(* IEC 61131-3 sources: dummvinci-rosetta-plc/src/plc_mcp/library/patterns, 6 files *)

(* ---- FB_AlarmManager.st ---- *)
(* =====================================================================
   FB_AlarmManager — aggregate N alarm points (IEC 62682 / ISA-18.2)
   dummvinci-rosetta-plc engineering library

   Aggregates the OUTPUT arrays of FB_AlarmPoint instances: per-class
   counts, unacked count, horn drive, and FIRST-OUT capture (which alarm
   started the trip cascade — the question every breakdown review asks).

   USAGE
     The application owns the FB_AlarmPoint instances and copies their
     outputs into the three arrays each cycle (or maps them directly):
       aActive[i]  := fbAlm_i.xActive;
       aUnacked[i] := fbAlm_i.xUnacked;
       aClass[i]   := fbAlm_i.eClass;
     then calls:
       fbMgr(nPoints := <used>, aActive := ..., aUnacked := ..., aClass := ...);
     Group acknowledge: wire fbMgr.xAckPulse into every point's xAck.
     Sizing: ARRAY[1..64] here — adjust bound + nPoints per project.

   DISCLAIMER — draft engineering input, review + FAT mandatory.
   NOT for safety-instrumented functions (SAFETY.md / H11).
   ===================================================================== *)

FUNCTION_BLOCK FB_AlarmManager
VAR_INPUT
    nPoints    : INT;    (* number of points actually used, <= 64 *)
    xGroupAck  : BOOL;   (* operator group-acknowledge command    *)
    xHornReset : BOOL;   (* silence horn without acknowledging    *)
END_VAR
VAR_IN_OUT
    aActive  : ARRAY[1..64] OF BOOL;
    aUnacked : ARRAY[1..64] OF BOOL;
    aClass   : ARRAY[1..64] OF INT;   (* 2 FAULT / 1 WARNING / 0 EVENT *)
END_VAR
VAR_OUTPUT
    nActive        : INT;
    nUnacked       : INT;
    nActiveFault   : INT;
    nActiveWarning : INT;
    iFirstOut      : INT;    (* index of first-out alarm, 0 = none *)
    xHorn          : BOOL;   (* unacked FAULT/WARNING present      *)
    xAckPulse      : BOOL;   (* wire into every point's xAck input *)
END_VAR
VAR
    i           : INT;
    aPrevActive : ARRAY[1..64] OF BOOL;
    nPrevActive : INT;
    xHornMuted  : BOOL;
    trigAck     : R_TRIG;
END_VAR

trigAck(CLK := xGroupAck);
xAckPulse := trigAck.Q;

nActive := 0;
nUnacked := 0;
nActiveFault := 0;
nActiveWarning := 0;

FOR i := 1 TO nPoints DO
    IF aActive[i] THEN
        nActive := nActive + 1;
        IF aClass[i] = 2 THEN
            nActiveFault := nActiveFault + 1;
        END_IF;
        IF aClass[i] = 1 THEN
            nActiveWarning := nActiveWarning + 1;
        END_IF;
    END_IF;
    IF aUnacked[i] THEN
        nUnacked := nUnacked + 1;
    END_IF;

    (* first-out: the point that went active while nothing was active *)
    IF aActive[i] AND NOT aPrevActive[i]
       AND (nPrevActive = 0) AND (iFirstOut = 0) THEN
        iFirstOut := i;
    END_IF;
    aPrevActive[i] := aActive[i];
END_FOR;

(* first-out clears only when the plant is alarm-free again *)
IF nActive = 0 THEN
    iFirstOut := 0;
END_IF;
nPrevActive := nActive;

(* horn: any unacked FAULT/WARNING; mute survives until all acked *)
IF xHornReset THEN
    xHornMuted := TRUE;
END_IF;
IF nUnacked = 0 THEN
    xHornMuted := FALSE;
END_IF;
xHorn := (nUnacked > 0) AND NOT xHornMuted;

END_FUNCTION_BLOCK

(* ---- FB_AlarmPoint.st ---- *)
(* =====================================================================
   FB_AlarmPoint — single alarm point state machine
   dummvinci-rosetta-plc engineering library

   STANDARD BASIS
     IEC 62682 / ISA-18.2 alarm states:
       0 = NORM        normal, inactive
       1 = UNACK_ALM   active, unacknowledged
       2 = ACK_ALM     active, acknowledged
       3 = UNACK_RTN   returned to normal, still unacknowledged
     Meldeklassen mapping (German practice):
       eClass 2 = FAULT   (Störung)   — trips/stops the function
       eClass 1 = WARNING (Warnung)   — degraded, action required
       eClass 0 = EVENT   (Meldung)   — information, logged only

   USAGE
     One instance per alarm point. Call every task cycle:
       fbAlm(xIn := <raw condition>, xAck := <ack cmd>, xReset := <reset>);
     Wire xAppeared/xDisappeared/xAckEdge into FB_EventLogger for the
     historian, and xActive/xUnacked/eClass arrays into FB_AlarmManager.

   DISCLAIMER — draft engineering input, review + FAT mandatory.
   NOT for safety-instrumented functions (see SAFETY.md / H11): e-stop,
   overload, interlock chains belong on a certified safety CPU.
   ===================================================================== *)

FUNCTION_BLOCK FB_AlarmPoint
VAR_INPUT
    xIn        : BOOL;   (* raw alarm condition, TRUE = abnormal *)
    xAck       : BOOL;   (* acknowledge command (operator/group)  *)
    xReset     : BOOL;   (* reset for latched alarms              *)
    xLatching  : BOOL;   (* TRUE: stays active until xReset       *)
    tOnDelay   : TIME;   (* debounce before alarm becomes active  *)
    tOffDelay  : TIME;   (* delay before return-to-normal         *)
    iPriority  : INT;    (* 1=low .. 4=critical (per philosophy)  *)
    eClass     : INT;    (* 2=FAULT, 1=WARNING, 0=EVENT           *)
    diCode     : DINT;   (* error code for catalog/historian      *)
END_VAR
VAR_OUTPUT
    xActive       : BOOL;  (* alarm condition present (qualified) *)
    xUnacked      : BOOL;  (* requires operator acknowledgement   *)
    eState        : INT;   (* 0 NORM / 1 UNACK_ALM / 2 ACK_ALM / 3 UNACK_RTN *)
    xAppeared     : BOOL;  (* one-cycle pulse: alarm appeared     *)
    xDisappeared  : BOOL;  (* one-cycle pulse: alarm cleared      *)
    xAckEdge      : BOOL;  (* one-cycle pulse: acknowledged       *)
END_VAR
VAR
    tonQualify  : TON;
    tonClear    : TON;
    xQualified  : BOOL;
    xLatched    : BOOL;
    trigApp     : R_TRIG;
    trigDis     : F_TRIG;
    trigAck     : R_TRIG;
END_VAR

(* --- qualification: debounce both directions ---------------------- *)
tonQualify(IN := xIn, PT := tOnDelay);
tonClear(IN := NOT xIn, PT := tOffDelay);

IF tonQualify.Q THEN
    xQualified := TRUE;
END_IF;
IF tonClear.Q THEN
    xQualified := FALSE;
END_IF;

(* --- latching ------------------------------------------------------ *)
IF xLatching AND xQualified THEN
    xLatched := TRUE;
END_IF;
IF xReset AND NOT xQualified THEN
    xLatched := FALSE;
END_IF;

xActive := xQualified OR (xLatching AND xLatched);

(* --- ack edge: evaluate BEFORE the state machine clears xUnacked --- *)
trigAck(CLK := xAck AND xUnacked);
xAckEdge := trigAck.Q;

(* --- IEC 62682 state machine --------------------------------------- *)
CASE eState OF
    0: (* NORM *)
        IF xActive THEN
            eState := 1;
            xUnacked := TRUE;
        END_IF;
    1: (* UNACK_ALM *)
        IF xAck THEN
            eState := 2;
            xUnacked := FALSE;
        ELSIF NOT xActive THEN
            eState := 3;
        END_IF;
    2: (* ACK_ALM *)
        IF NOT xActive THEN
            eState := 0;
        END_IF;
    3: (* UNACK_RTN *)
        IF xAck THEN
            eState := 0;
            xUnacked := FALSE;
        ELSIF xActive THEN
            eState := 1;
        END_IF;
END_CASE;

(* --- edges for the historian ---------------------------------------- *)
trigApp(CLK := xActive);
xAppeared := trigApp.Q;
trigDis(CLK := xActive);
xDisappeared := trigDis.Q;

END_FUNCTION_BLOCK

(* ---- FB_CommsWatchdog.st ---- *)
(* =====================================================================
   FB_CommsWatchdog — communication supervision (DIAGNOSTICS ONLY)
   dummvinci-rosetta-plc engineering library

   Supervises a cyclic link (Modbus TCP slave, HMI, remote I/O) via a
   heartbeat counter that the remote increments. If the counter stops
   changing for tTimeout, the link is declared down — feed that into an
   FB_AlarmPoint (class WARNING or FAULT per the alarm philosophy).

   ⚠ THIS IS NOT A SAFETY WATCHDOG. A watchdog whose timeout must bring
   the machine to a safe state is a safety function — that belongs on a
   certified safety CPU (AC500-S) per SAFETY.md / hazard H11. This block
   only *reports* link health.

   USAGE (Modbus TCP to an ACS880 example)
     Map a drive register that changes continuously (e.g. a counter or
     the actual-speed word) into diHeartbeat:
       fbWd(diHeartbeat := <mapped register>, tTimeout := T#3s);

   DISCLAIMER — draft engineering input, review + FAT mandatory.
   ===================================================================== *)

FUNCTION_BLOCK FB_CommsWatchdog
VAR_INPUT
    diHeartbeat : DINT;   (* value the remote updates cyclically *)
    tTimeout    : TIME;   (* declare down after this long unchanged *)
END_VAR
VAR_OUTPUT
    xCommsOk  : BOOL;
    xTimeout  : BOOL;
    udiDrops  : UDINT;    (* number of times the link went down *)
END_VAR
VAR
    diPrev   : DINT;
    tonStale : TON;
    trigDown : R_TRIG;
END_VAR

tonStale(IN := (diHeartbeat = diPrev), PT := tTimeout);
diPrev := diHeartbeat;

xTimeout := tonStale.Q;
xCommsOk := NOT xTimeout;

trigDown(CLK := xTimeout);
IF trigDown.Q THEN
    udiDrops := udiDrops + 1;
END_IF;

END_FUNCTION_BLOCK

(* ---- FB_DriveDiagACS880.st ---- *)
(* =====================================================================
   FB_DriveDiagACS880 — ACS880 fault/warning capture for the historian
   dummvinci-rosetta-plc engineering library

   Captures the active fault/warning codes of an ABB ACS880 drive (read
   over Modbus TCP / PROFINET) and converts them to hex strings that key
   directly into the error-code catalog (plc_errorcode_lookup, source
   "acs880") for cause + remedy.

   REGISTER MAPPING (project-specific — TODO verify against YOUR comms
   mapping in Drive Composer Pro; typical parameters):
     04.01  Tripping fault code    -> uiFaultCode
     04.06  Active warning code    -> uiWarnCode
     Status word bit FAULTED       -> xDriveFaulted
     Status word bit WARNING       -> xDriveWarning

   USAGE
     fbDiag(uiFaultCode := <mapped 04.01>, uiWarnCode := <mapped 04.06>,
            xDriveFaulted := <SW bit>, xDriveWarning := <SW bit>);
     On xNewFault: log to FB_EventLogger with diCode := fbDiag.diFaultCode
     and look the hex string up in the catalog.

   DISCLAIMER — draft engineering input, review + FAT mandatory. Codes and
   remedies come from the catalog, which must be verified against the
   ACS880 firmware manual for the installed FW revision.
   ===================================================================== *)

FUNCTION_BLOCK FB_DriveDiagACS880
VAR_INPUT
    uiFaultCode   : UINT;   (* drive par 04.01 via comms *)
    uiWarnCode    : UINT;   (* drive par 04.06 via comms *)
    xDriveFaulted : BOOL;   (* status word: faulted      *)
    xDriveWarning : BOOL;   (* status word: warning      *)
END_VAR
VAR_OUTPUT
    xFault      : BOOL;
    xWarning    : BOOL;
    diFaultCode : DINT;         (* numeric, for FB_EventLogger *)
    sFaultHex   : STRING(7);    (* catalog key, e.g. '2310'    *)
    sWarnHex    : STRING(7);
    xNewFault   : BOOL;         (* one-cycle pulse             *)
    xNewWarning : BOOL;
END_VAR
VAR
    trigF : R_TRIG;
    trigW : R_TRIG;
    uiTmp : UINT;
    iNib  : INT;
    i     : INT;
    sHex  : STRING(7);
END_VAR

xFault := xDriveFaulted;
xWarning := xDriveWarning;
diFaultCode := TO_DINT(uiFaultCode);

(* --- UINT -> 4-digit hex string (ACS880 codes read as hex) ---------
   MID signature per IEC 61131-3 / CODESYS Standard library:
   MID(IN, L, P) = L characters starting at position P (1-based).
   So MID('0123456789ABCDEF', L := 1, P := iNib + 1) extracts exactly
   ONE nibble character. Do not swap to (pos, len) — that is a
   different vendor convention. ------------------------------------- *)
sHex := '';
uiTmp := uiFaultCode;
FOR i := 1 TO 4 DO
    iNib := TO_INT(uiTmp MOD 16);
    sHex := CONCAT(MID(IN := '0123456789ABCDEF', L := 1, P := iNib + 1),
                   sHex);
    uiTmp := uiTmp / 16;
END_FOR;
sFaultHex := sHex;

sHex := '';
uiTmp := uiWarnCode;
FOR i := 1 TO 4 DO
    iNib := TO_INT(uiTmp MOD 16);
    sHex := CONCAT(MID(IN := '0123456789ABCDEF', L := 1, P := iNib + 1),
                   sHex);
    uiTmp := uiTmp / 16;
END_FOR;
sWarnHex := sHex;

trigF(CLK := xDriveFaulted);
xNewFault := trigF.Q;
trigW(CLK := xDriveWarning);
xNewWarning := trigW.Q;

END_FUNCTION_BLOCK

(* ---- FB_EventLogger.st ---- *)
(* =====================================================================
   FB_EventLogger — sequence-of-events ring-buffer historian
   dummvinci-rosetta-plc engineering library

   In-PLC SoE log: every alarm appearance/clearance/acknowledgement is
   stamped and kept in a retained ring buffer for breakdown analysis and
   HMI display. Design rationale: docs/library/HISTORIAN-DESIGN.md
   (resolution limits, time sync, when to use an external historian).

   USAGE
     One instance per log. Feed one event per rising edge of xLog —
     typically chained from FB_AlarmPoint edges:
       IF fbAlm.xAppeared THEN
           fbLog(xLog := TRUE, diCode := fbAlm.diCode,
                 eClass := fbAlm.eClass, eEdge := 0, rValue := <pv>,
                 dtNow := <rtc>, uiMsOfSec := <ms>);
       END_IF
     eEdge: 0 = APPEARED, 1 = DISAPPEARED, 2 = ACKED.
     (* TODO platform binding: dtNow/uiMsOfSec must come from the CPU RTC
        — e.g. AC500 V3 SysTimeRtc / DT clock FBs. Timestamp AT SOURCE,
        in the same task that detects the edge. *)
     Buffer: ARRAY[0..255] here — size per project; RETAIN memory is a
     real CPU budget, verify against the CPU's retain capacity.

   TYPES (move to a DUT object on Automation Builder import)
   ===================================================================== *)

TYPE ST_Event :
STRUCT
    udiSeq     : UDINT;   (* monotonic sequence number         *)
    dtStamp    : DT;      (* RTC date-time                     *)
    uiMs       : UINT;    (* millisecond-of-second, if available *)
    diCode     : DINT;    (* error/alarm code (catalog key)    *)
    eClass     : INT;     (* 2 FAULT / 1 WARNING / 0 EVENT     *)
    eEdge      : INT;     (* 0 APPEARED / 1 DISAPPEARED / 2 ACKED *)
    rValue     : REAL;    (* process value at event time       *)
END_STRUCT
END_TYPE

FUNCTION_BLOCK FB_EventLogger
VAR_INPUT
    xLog       : BOOL;    (* rising edge stores one event  *)
    dtNow      : DT;      (* TODO platform: bind to CPU RTC *)
    uiMsOfSec  : UINT;
    diCode     : DINT;
    eClass     : INT;
    eEdge      : INT;
    rValue     : REAL;
END_VAR
VAR_OUTPUT
    uiHead     : UINT;    (* index of most recent event    *)
    udiTotal   : UDINT;   (* events logged since power-up of retain *)
    xWrapped   : BOOL;    (* buffer has overwritten old entries *)
END_VAR
VAR
    trigLog : R_TRIG;
END_VAR
VAR RETAIN
    aBuf   : ARRAY[0..255] OF ST_Event;
    uiNext : UINT;
    udiSeq : UDINT;
END_VAR

trigLog(CLK := xLog);
IF trigLog.Q THEN
    aBuf[uiNext].udiSeq  := udiSeq;
    aBuf[uiNext].dtStamp := dtNow;
    aBuf[uiNext].uiMs    := uiMsOfSec;
    aBuf[uiNext].diCode  := diCode;
    aBuf[uiNext].eClass  := eClass;
    aBuf[uiNext].eEdge   := eEdge;
    aBuf[uiNext].rValue  := rValue;
    uiHead := uiNext;
    uiNext := (uiNext + 1) MOD 256;
    udiSeq := udiSeq + 1;
    udiTotal := udiSeq;
    IF udiSeq > 256 THEN
        xWrapped := TRUE;
    END_IF;
END_IF;

END_FUNCTION_BLOCK

(* ---- FB_FaultLatch.st ---- *)
(* =====================================================================
   FB_FaultLatch — lightweight fault latch with shared first-out capture
   dummvinci-rosetta-plc engineering library

   For simple trip chains where the full FB_AlarmPoint state machine is
   overkill: latch on fault, hold until reset, and capture whether THIS
   fault was the first of the cascade (shared group flag).

   USAGE
     One shared BOOL per fault group:
       VAR xGrpFirstOutTaken : BOOL; END_VAR
     Per fault:
       fbFault(xIn := <condition>, xReset := <reset cmd>,
               xGroupFirstOutTaken := xGrpFirstOutTaken);
     The application clears xGrpFirstOutTaken when the group is healthy
     again (all xLatched FALSE).

   DISCLAIMER — draft engineering input, review + FAT mandatory.
   NOT for safety-instrumented functions (SAFETY.md / H11).
   ===================================================================== *)

FUNCTION_BLOCK FB_FaultLatch
VAR_INPUT
    xIn    : BOOL;   (* fault condition, TRUE = faulted *)
    xReset : BOOL;   (* reset command                   *)
END_VAR
VAR_IN_OUT
    xGroupFirstOutTaken : BOOL;   (* shared across the fault group *)
END_VAR
VAR_OUTPUT
    xLatched  : BOOL;
    xFirstOut : BOOL;   (* TRUE if this fault started the cascade *)
END_VAR

IF xIn THEN
    IF NOT xLatched AND NOT xGroupFirstOutTaken THEN
        xFirstOut := TRUE;
        xGroupFirstOutTaken := TRUE;
    END_IF;
    xLatched := TRUE;
END_IF;

IF xReset AND NOT xIn THEN
    xLatched := FALSE;
    xFirstOut := FALSE;
END_IF;

END_FUNCTION_BLOCK
